(*
	Exporter test double that captures the linked list a processor transfers via
	export, so tests can assert on the exported batch. Set busy to
	simulate an exporter that cannot accept a batch. callsWhileBusy counts
	export calls made while busy, which a processor must never make.
*)
FUNCTION_BLOCK FB_LogRecordExporter_ForInspection EXTENDS FB_LogRecordExporter_Base
VAR_INPUT
	busy: BOOL;		// TRUE simulates a busy exporter that refuses batches
END_VAR
VAR_OUTPUT
	callsWhileBusy: UDINT;
END_VAR

METHOD isBusy : BOOL
isBusy := THIS^.busy;
END_METHOD

// the captured batch, for test assertions
PROPERTY records : REFERENCE TO FB_LogRecordQueue
GET
records REF= THIS^._records;
END_GET
END_PROPERTY

METHOD tick : BOOL
VAR_OUTPUT
	failureReason: E_LogRecordExporterFailureReason;
END_VAR
failureReason := E_LogRecordExporterFailureReason.NA;
tick := TRUE;
END_METHOD

METHOD export : BOOL
VAR_IN_OUT
	logRecords: FB_LogRecordQueue;
END_VAR
VAR_INPUT
	count: UDINT;
END_VAR
VAR_OUTPUT
	failureReason: E_LogRecordExporterFailureReason;
END_VAR
IF THIS^.isBusy() THEN
	THIS^.callsWhileBusy := THIS^.callsWhileBusy + 1;
END_IF
export := SUPER^.export(logRecords:=logRecords, count:=count, failureReason=>failureReason);
END_METHOD

END_FUNCTION_BLOCK

(* stored: Version 1.1.0.1
   POU FB_LogRecordExporter_ForInspection: Id {d4b9a2e7-6f31-48c5-9b0a-1e8c72d5f4a3}, SpecialFunc None
   Method isBusy: Id {a1f83d64-92b7-4e5a-8c39-7d15b0e6c2f9}
   Property records: Id {3c6e94b1-58d2-4f7a-a0e4-2b91c8d5a7f6}
   Get Get: Id {6b28d5f3-1c97-4e40-b8a2-5f04e9c3d1a8}
   Method tick: Id {900e1bfc-7fef-4279-8923-fb8a822cc1c3}
   Method export: Id {e330627d-8bfe-470b-94c7-55d6e8d5acfc} *)
